FUNCTION_BLOCK IO_DO (* One digital output (a motor's enable, a direction, a valve). Its Address says where the signal goes: a Raspberry Pi pin, a Modbus coil, or simulated. Technical: Digital output; Address: 'gpio[chip:line(:pull_up|:pull_down)(:active_low)]' or 'pwm[chip:channel:period_ns]' a Raspberry Pi's line, set up here; 'modbus[...]' a Modbus CLIENT ID; 'sim' simulated; another name a local IO handle set up elsewhere (QX PARAMS); empty: not connected (QO = FALSE) *)
  (* Standard: 61499-2 *)
  (* Version 0.1, 2026-09-28, Project contributors, AAU Smart Production Lab *)
  PACKAGE modlib;
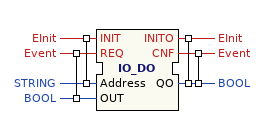
  EVENT_INPUT
    INIT : EInit WITH Address; (* Set up the point from Address (at start-up) *)
    REQ WITH OUT; (* Read the point, or write OUT to it *)
  END_EVENT
  EVENT_OUTPUT
    INITO : EInit WITH QO; (* Set up: QO says whether the point is reachable *)
    CNF WITH QO; (* Done: QO says whether it worked (an input: IN is the value read) *)
  END_EVENT
  VAR_INPUT
    Address : STRING; (* Where the point is: 'gpio[chip:line(:pull_up|:pull_down)(:active_low)]', 'pwm[chip:channel:period_ns]', 'modbus[...]', 'sim', or an IO handle's name; empty: not connected *)
    OUT : BOOL; (* The value to write *)
  END_VAR
  VAR_OUTPUT
    QO : BOOL; (* The point is reachable, the last access worked *)
  END_VAR
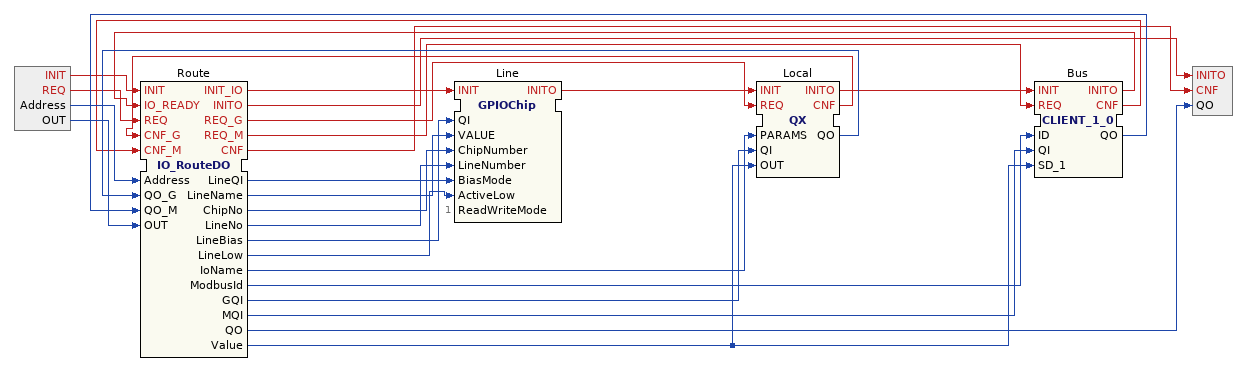
  FBS
    Route : modlib::IO_RouteDO; (* Picks the way to the signal from the Address and passes values that way. *)
    Line : eclipse4diac::io::gpiochip::GPIOChip(ReadWriteMode := 1); (* Sets up a Raspberry Pi line (GPIO) or PWM channel when the Address names one. *)
    Local : eclipse4diac::io::QX; (* Reads or writes a FORTE IO handle (IX, QX, IW, QW). *)
    Bus : iec61499::net::CLIENT_1_0; (* Reads or writes a Modbus register when the Address names one. *)
  END_FBS
  EVENT_CONNECTIONS
    INIT TO Route.INIT;
    Route.INIT_IO TO Line.INIT;
    Line.INITO TO Local.INIT;
    Local.INITO TO Bus.INIT;
    Bus.INITO TO Route.IO_READY;
    Route.INITO TO INITO;
    REQ TO Route.REQ;
    Route.REQ_G TO Local.REQ;
    Route.REQ_M TO Bus.REQ;
    Local.CNF TO Route.CNF_G;
    Bus.CNF TO Route.CNF_M;
    Route.CNF TO CNF;
  END_CONNECTIONS
  DATA_CONNECTIONS
    Route.LineQI TO Line.QI;
    Route.LineName TO Line.VALUE;
    Route.ChipNo TO Line.ChipNumber;
    Route.LineNo TO Line.LineNumber;
    Route.LineBias TO Line.BiasMode;
    Route.LineLow TO Line.ActiveLow;
    Address TO Route.Address;
    Route.IoName TO Local.PARAMS;
    Route.ModbusId TO Bus.ID;
    Route.GQI TO Local.QI;
    Route.MQI TO Bus.QI;
    Local.QO TO Route.QO_G;
    Bus.QO TO Route.QO_M;
    Route.QO TO QO;
    OUT TO Route.OUT;
    Route.Value TO Local.OUT;
    Route.Value TO Bus.SD_1;
  END_CONNECTIONS
END_FUNCTION_BLOCK
